SUBAPPLICATION GreenWhiteRedBackground3_AX (* Hintergrundfarbe fuer SoftKey + Aux (3 Objekte), 3 Zustaende: DI1 FALSE -> Weiss, TRUE -> Gruen, DI2 TRUE -> Rot (Vorrang) *)
  (* Standard: 61499-2; Description: Copyright (c) 2026 Meisterschulen am Ostbahnhof This program and the accompanying materials are made available under the terms of the Eclipse Public License 2.0 which is available at https://www.eclipse.org/legal/epl-2.0/ SPDX-License-Identifier: EPL-2.0 *)
  (* Version 1.0, 2026-10-29, Franz Höpfinger, Meisterschulen am Ostbahnhof, Neu, Muster WhiteGreenPurpleBackground1_AX (AUS-Adapter-Kette), Objekte wie GreenWhiteBackground3_AX. Franz: GreenWhiteRed mit 2x AX, ROT hat Vorrang vor GRUEN. Gedacht fuer DI2 = Station nicht erreichbar. *)
  PACKAGE MyLib::sys;
  IMPORT isobus::UT::Q::const::IDs::ID_NULL;
  IMPORT isobus::UT::Q::const::colours::COLOR_GREEN;
  IMPORT isobus::UT::Q::const::colours::COLOR_WHITE;
  IMPORT isobus::UT::Q::const::colours::COLOR_RED;
  (* Documentation:
  Hintergrundfarbe Grün/Weiß/Rot für SoftKey + Aux
   Wie GreenWhiteBackground3_AX (DI1: TRUE → Grün, FALSE → Weiß, für SoftKey, Aux-Vorschau und Aux-Handle), zusätzlich DI2: TRUE → Rot, mit Vorrang vor DI1. Aufbau wie WhiteGreenPurpleBackground1_AX (AUS-Adapter-Kette, jede Änderung von DI1 oder DI2 liefert die vollständige Farbe).
   Einsatz: DI2 = Station nicht erreichbar (invertiertes ALIVE aus Station_Alive_VT_OPC), damit die Taste keinen veralteten Zustand zeigt.
  *)
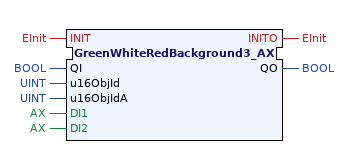
  EVENT_INPUT
    INIT : EInit; (* Initialization Request *)
  END_EVENT
  EVENT_OUTPUT
    INITO : EInit; (* Initialization Confirm *)
  END_EVENT
  VAR_INPUT
    QI : BOOL := TRUE; (* Quality Input - TRUE to enable service *)
    u16ObjId : UINT := ID_NULL; (* Object ID Softkey *)
    u16ObjIdA : UINT := ID_NULL; (* Object ID AUX *)
  END_VAR
  VAR_OUTPUT
    QO : BOOL; (* Quality Output - TRUE if service executed successfully (AND aller Instanzen) *)
  END_VAR
  SOCKETS
    DI1 : adapter::types::unidirectional::AX; (* Zustand (FALSE=Weiss, TRUE=Gruen) *)
    DI2 : adapter::types::unidirectional::AX; (* TRUE=Rot, Vorrang vor DI1 *)
  END_SOCKETS
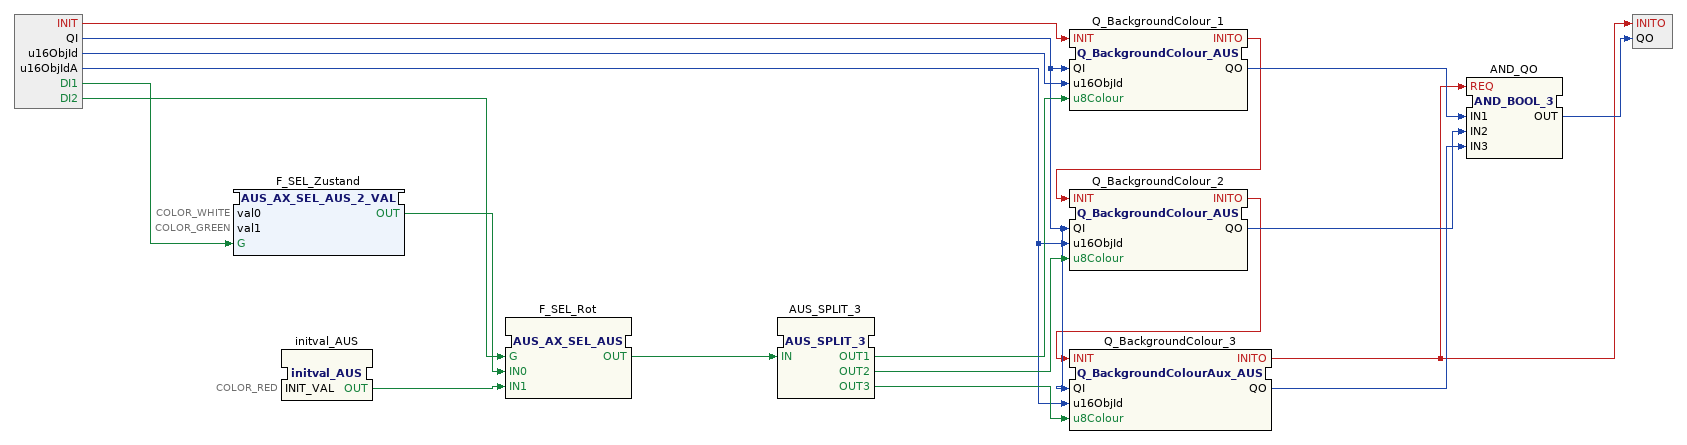
  FBS
    F_SEL_Rot : adapter::iec61131::selection::AUS_AX_SEL_AUS;
    initval_AUS : adapter::types::unidirectional::AUS::initval::initval_AUS(INIT_VAL := COLOR_RED);
    AUS_SPLIT_3 : adapter::events::unidirectional::AUS_SPLIT_3;
    Q_BackgroundColour_1 : isobus::UT::Q::Q_BackgroundColour_AUS;
    Q_BackgroundColour_2 : isobus::UT::Q::Q_BackgroundColour_AUS;
    Q_BackgroundColour_3 : isobus::UT::Q::Q_BackgroundColourAux_AUS;
    AND_QO : iec61131::booleanOperators::AND_BOOL_3;
  END_FBS
  SUBAPPS
    F_SEL_Zustand : MyLib::sys::AUS_AX_SEL_AUS_2_VAL(val0 := COLOR_WHITE, val1 := COLOR_GREEN);
  END_SUBAPPS
  EVENT_CONNECTIONS
    INIT TO Q_BackgroundColour_1.INIT;
    Q_BackgroundColour_1.INITO TO Q_BackgroundColour_2.INIT;
    Q_BackgroundColour_2.INITO TO Q_BackgroundColour_3.INIT;
    Q_BackgroundColour_3.INITO TO AND_QO.REQ;
    Q_BackgroundColour_3.INITO TO INITO;
  END_CONNECTIONS
  DATA_CONNECTIONS
    QI TO Q_BackgroundColour_1.QI;
    QI TO Q_BackgroundColour_2.QI;
    QI TO Q_BackgroundColour_3.QI;
    u16ObjId TO Q_BackgroundColour_1.u16ObjId;
    u16ObjIdA TO Q_BackgroundColour_2.u16ObjId;
    u16ObjIdA TO Q_BackgroundColour_3.u16ObjId;
    Q_BackgroundColour_1.QO TO AND_QO.IN1;
    Q_BackgroundColour_2.QO TO AND_QO.IN2;
    Q_BackgroundColour_3.QO TO AND_QO.IN3;
    AND_QO.OUT TO QO;
  END_CONNECTIONS
  ADAPTER_CONNECTIONS
    DI1 TO F_SEL_Zustand.G;
    DI2 TO F_SEL_Rot.G;
    F_SEL_Zustand.OUT TO F_SEL_Rot.IN0;
    initval_AUS.OUT TO F_SEL_Rot.IN1;
    F_SEL_Rot.OUT TO AUS_SPLIT_3.IN;
    AUS_SPLIT_3.OUT1 TO Q_BackgroundColour_1.u8Colour;
    AUS_SPLIT_3.OUT2 TO Q_BackgroundColour_2.u8Colour;
    AUS_SPLIT_3.OUT3 TO Q_BackgroundColour_3.u8Colour;
  END_CONNECTIONS
END_SUBAPPLICATION
